Universal Robots PolyScope program: rg2.urp

Program rg2 (installation=default directory=/programs/new folder createdIn=5.11.11.1010533 lastSavedIn=5.11.11.1010533 robotSerialNumber=20195501451)
Calibrated DH parameters: a=[0.000053, -0.349069, -0.379258, 0.00007, -0.000011, 0]; d=[0.162389, 188.384002, -210.84231, 22.591517, 0.099817, 0.099561]; alpha=[1.570074, -0.001289, -0.004473, 1.570456, -1.569854, 0]; deltaTheta=[0, -0.607882, 7.150013, -0.258941, 0, 0]
Robot Program (runOnlyOnce=false)
  URCap RG2 (RG - On Robot, OnRobot A/S) dataModel(depthCompensate=false, width=0, force=40, payload=0.0, name=RG2(0))
